// TIA Portal V21 export
// export: Created 2026-11-21T10:55:36.0058378Z, ExportSetting WithDefaults, DisplayName Totally Integrated Automation Portal, DisplayVersion V21, DisplayName STEP 7 Professional, DisplayVersion V21, DisplayName STEP 7 Safety, DisplayVersion V21, DisplayName Tech WebApplication, DisplayVersion V21, DisplayName WinCC Basic/Comfort/Advanced, DisplayVersion V21, DisplayName WinCC Unified, DisplayVersion V21
VAR_GLOBAL   // PLC tag table "Inputs"
   Button_Start AT %I0.0 : Bool;   // Start the line
   Button_Stop AT %I0.1 : Bool;   // Stop the line, normally closed
   Button_Reset AT %I0.2 : Bool;   // Acknowledge faults
   Infeed_BottleAtFiller AT %I1.0 : Bool;   // Photo eye: a bottle stands under the filler
   Infeed_MotorFeedback AT %I1.1 : Bool;   // Infeed contactor is closed
   Outfeed_BottleAtEnd AT %I1.2 : Bool;   // Photo eye at the end of the outfeed
   Outfeed_MotorFeedback AT %I1.3 : Bool;   // Outfeed contactor is closed
   Filler_ValveOpened AT %I1.4 : Bool;   // Fill valve is open
   Filler_ValveClosed AT %I1.5 : Bool;   // Fill valve is closed
   Packer_Ready AT %I1.6 : Bool;   // The packer can take a bottle
   Filler_Level AT %IW64 : Int;   // Level in the bottle, raw 0 to 27648
END_VAR
